(* IEC 61131-3 sources: axsharp/src/ix.compiler/tests/Ix.Compiler.CsTests/samples/units/src, 32 files *)

(* ---- compileromitsattribute.st ---- *)
NAMESPACE CompilerOmmits
    CLASS ClassWithArrays
        VAR PUBLIC
            {#ix-attr:[CompilerOmitsAttribute()]}
            _must_be_omitted_everywhere : Complex;
            {#ix-attr:[CompilerOmitsAttribute("Onliner")]}
            _must_be_omitted_in_onliner : Complex;
            {#ix-attr:[CompilerOmitsAttribute("POCO")]}
             _must_be_omitted_in_poco : Complex;
            _primitive  : ARRAY[0..10] OF BYTE;
        END_VAR

    END_CLASS

    CLASS PUBLIC Complex
        VAR PUBLIC
            HelloString : STRING;
            Id : ULINT;
        END_VAR
    END_CLASS
END_NAMESPACE

NAMESPACE Enums
    CLASS ClassWithEnums
        VAR PUBLIC
            colors : Colors;
            NamedValuesColors : NamedValuesColors;
        END_VAR

    END_CLASS

    TYPE
        Colors : (Red, Green, Blue) := Red;
    END_TYPE

    TYPE
        NamedValuesColors : STRING (Red := '1', Green := '2', Blue := '3') := Red;
    END_TYPE

END_NAMESPACE

NAMESPACE misc
    CLASS PUBLIC VariousMembers
        VAR PUBLIC
            _SomeClass : SomeClass;
            _Motor : Motor;
        END_VAR
    END_CLASS

    CLASS SomeClass
        VAR PUBLIC
            SomeClassVariable : STRING;
        END_VAR
    END_CLASS

    TYPE
        Motor : STRUCT
            isRunning : BOOL;
        END_STRUCT;
        Vehicle : STRUCT
            m : Motor;
            displacement : INT;
        END_STRUCT;
    END_TYPE
END_NAMESPACE

NAMESPACE UnknownArraysShouldNotBeTraspiled
    CLASS ClassWithArrays
        VAR PUBLIC
            _complexKnown : ARRAY[0..10] OF Complex;
            _complexUnknown : ARRAY [0..10] OF ComplexUnknown;
            _primitive  : ARRAY[0..10] OF BYTE;
        END_VAR

    END_CLASS

    CLASS PUBLIC Complex
        VAR PUBLIC
            HelloString : STRING;
            Id : ULINT;
        END_VAR
    END_CLASS
END_NAMESPACE

(* ---- enum_simple.st ---- *)
TYPE
    Colors : (Red, Green, Blue) := Red;
END_TYPE

(* ---- misc.st ---- *)
NAMESPACE Enums
    CLASS ClassWithEnums
        VAR PUBLIC
            colors : Colors;
            NamedValuesColors : NamedValuesColors;
        END_VAR

    END_CLASS

    TYPE
        Colors : (Red, Green, Blue) := Red;
    END_TYPE

    TYPE
        NamedValuesColors : STRING (Red := '1', Green := '2', Blue := '3') := Red;
    END_TYPE

END_NAMESPACE

NAMESPACE misc
    CLASS PUBLIC VariousMembers
        VAR PUBLIC
            _SomeClass : SomeClass;
            _Motor : Motor;
        END_VAR
    END_CLASS

    CLASS SomeClass
        VAR PUBLIC
            SomeClassVariable : STRING;
        END_VAR
    END_CLASS

    TYPE
        Motor : STRUCT
            isRunning : BOOL;
        END_STRUCT;
        Vehicle : STRUCT
            m : Motor;
            displacement : INT;
        END_STRUCT;
    END_TYPE
END_NAMESPACE

NAMESPACE UnknownArraysShouldNotBeTraspiled
    CLASS ClassWithArrays
        VAR PUBLIC
            _complexKnown : ARRAY[0..10] OF Complex;
            _complexUnknown : ARRAY [0..10] OF ComplexUnknown;
            _primitive  : ARRAY[0..10] OF BYTE;
        END_VAR

    END_CLASS

    CLASS PUBLIC Complex
        VAR PUBLIC
            HelloString : STRING;
            Id : ULINT;
        END_VAR
    END_CLASS
END_NAMESPACE

(* ---- struct_simple.st ---- *)
TYPE
    Motor : STRUCT
        isRunning : BOOL;
    END_STRUCT;
    Vehicle : STRUCT
        m : Motor;
        displacement : INT;
    END_STRUCT;
END_TYPE

(* ---- type_named_values.st ---- *)
NAMESPACE NamedValuesNamespace
    TYPE
        LightColors : INT (
            LRED := 12,
            LGREEN := 14,
            LBLUE := 23
        );
    END_TYPE

    CLASS PUBLIC using_type_named_values
        VAR PUBLIC
            LColors : LightColors;
        END_VAR
    END_CLASS
END_NAMESPACE

(* ---- type_named_values_literals.st ---- *)
NAMESPACE Simatic.Ax.StateFramework
    TYPE
        StateControllerStatus : WORD (
            STATUS_NO_ERR := WORD#16#7000,
            STATUS_IS_RUNNING := WORD#16#7001,
            STATUS_STATE_CHANGED := WORD#16#7002,
            STATUS_NO_INITIALSTATE := WORD#16#8100,
            STATUS_NO_NEXTSTATE := WORD#16#8101
        ) := STATUS_NO_ERR;
    END_TYPE

    CLASS PUBLIC using_type_named_values
        VAR PUBLIC
            LColors : StateControllerStatus;
        END_VAR
    END_CLASS
END_NAMESPACE

(* ---- type_with_enum.st ---- *)
NAMESPACE Simatic.Ax.StateFramework
    INTERFACE IGuard

        METHOD Check : BOOL
        END_METHOD

        METHOD Reset
        END_METHOD

    END_INTERFACE
END_NAMESPACE

NAMESPACE Simatic.Ax.StateFramework

    /// Condition
    /// GT: Greater than compareValue
    /// EQ: Equal to compareValue
    /// LT: Less than compareValue
    /// NE: Is not equal to compareValue
    /// GE: Greater or equal to compareValue
    /// LE: Less or equal to compareValue
    TYPE
        Condition : (GT, EQ, LT, NE, GE, LE);
    END_TYPE

    CLASS CompareGuardLint IMPLEMENTS IGuard
        VAR PUBLIC
            Value : REF_TO LINT;
            CompareToValue : LINT;
            Condition : Condition;
        END_VAR

        METHOD PUBLIC Config
            VAR_INPUT
                countValue : REF_TO LINT;
                compareValue : LINT;
                compareCondition : Condition;
            END_VAR
            Value := countValue;
            CompareToValue := compareValue;
            Condition := compareCondition;
        END_METHOD

        // ---------------- IMPLEMENT IGuard---------------------------
        METHOD PUBLIC Check : BOOL

            CASE Condition OF
                Condition#GT : Check := Value^ > CompareToValue;
                Condition#EQ : Check := Value^ = CompareToValue;
                Condition#LT : Check := Value^ < CompareToValue;
                Condition#GE : Check := Value^ >= CompareToValue;
                Condition#LE : Check := Value^ <= CompareToValue;
            END_CASE
            ;

        END_METHOD

        METHOD PUBLIC Reset
            ;
        END_METHOD
        // ---------------- END IMPLEMENT IGuard---------------------------

    END_CLASS
END_NAMESPACE

(* ---- types_with_name_attributes.st ---- *)
NAMESPACE TypeWithNameAttributes
    TYPE
        {#ix-attr:[Container(Layout.Wrap)]}
        Motor : STRUCT
            isRunning : BOOL;
        END_STRUCT;
        Vehicle : STRUCT
            m : Motor;
            displacement : INT;
        END_STRUCT;
    END_TYPE

    {#ix-prop:public string AttributeName}
    CLASS NoAccessModifierClass
        VAR PUBLIC
            SomeClassVariable : STRING;
        END_VAR
    END_CLASS
END_NAMESPACE

(* ---- class_extends_and_implements.st ---- *)
CLASS PUBLIC ExtendsAndImplements EXTENDS ExtendeeExtendsAndImplements IMPLEMENTS IImplementation1, IImplementation2

END_CLASS

CLASS PUBLIC ExtendeeExtendsAndImplements

END_CLASS

INTERFACE PUBLIC IImplementation1 END_INTERFACE
INTERFACE PUBLIC IImplementation2 END_INTERFACE

(* ---- class_implements.st ---- *)
CLASS PUBLIC _NULL_CONTEXT IMPLEMENTS IContext

END_CLASS

INTERFACE PUBLIC IContext

END_INTERFACE

(* ---- class_implements_multiple.st ---- *)
CLASS PUBLIC _NULL_CONTEXT_MULTIPLE IMPLEMENTS IContext_Multiple, IObject_Multiple

END_CLASS

INTERFACE PUBLIC IContext_Multiple

END_INTERFACE

INTERFACE PUBLIC IObject_Multiple

END_INTERFACE

(* ---- file_with_unsupported.st ---- *)
NAMESPACE Unsupported
  FUNCTION SomeFunction : INT
    ;
  END_FUNCTION
END_NAMESPACE

(* ---- array_declaration.st ---- *)
NAMESPACE ArrayDeclarationSimpleNamespace
    CLASS array_declaration_class
        VAR PUBLIC
            primitive : ARRAY[1..100] OF INT;
            complex : ARRAY[1..100] OF some_complex_type;
        END_VAR
    END_CLASS

    CLASS some_complex_type
        VAR

        END_VAR

    END_CLASS

END_NAMESPACE

(* ---- class_all_primitives.st ---- *)
CLASS class_all_primitives
    VAR PUBLIC
        myBOOL	        :       BOOL	      ;
        myBYTE	        :       BYTE	      ;
        myWORD	        :       WORD	      ;
        myDWORD	        :       DWORD	      ;
        myLWORD	        :       LWORD	      ;
        mySINT	        :       SINT	      ;
        myINT	        :       INT	          ;
        myDINT	        :       DINT	      ;
        myLINT	        :       LINT	      ;
        myUSINT	        :       USINT	      ;
        myUINT	        :       UINT	      ;
        myUDINT	        :       UDINT	      ;
        myULINT	        :       ULINT	      ;
        myREAL	        :       REAL	      ;
        myLREAL	        :       LREAL	      ;
        myTIME	        :       TIME	      ;
        myLTIME	        :       LTIME	      ;
        myDATE	        :       DATE	      ;
     //   myLDATE	        :       LDATE	      ;
        myTIME_OF_DAY	:       TIME_OF_DAY	  ;
     //   myLTIME_OF_DAY	:       LTIME_OF_DAY  ;
        myDATE_AND_TIME  :      DATE_AND_TIME ;
     //   myLDATE_AND_TIME :      LDATE_AND_TIME;
     //   myCHAR	        :       CHAR	      ;
     //   myWCHAR	        :       WCHAR	      ;
        mySTRING	        :   STRING	      ;
        myWSTRING	    :       WSTRING	      ;
    END_VAR
END_CLASS

(* ---- class_extended_by_known_type.st ---- *)
USING Simatic.Ax.Stateframework;
USING Simatic.Ax.StatePattern;

NAMESPACE Simatic.Ax.StateFramework
    CLASS State1Transition EXTENDS AbstractState

        METHOD PUBLIC OVERRIDE OnEntry
            ;
        END_METHOD

        METHOD PUBLIC OVERRIDE OnExit
            ;
        END_METHOD

        METHOD PUBLIC OVERRIDE Action
            ;
        END_METHOD

    END_CLASS

END_NAMESPACE

NAMESPACE Simatic.Ax.StateFramework
    CLASS ABSTRACT AbstractState IMPLEMENTS IState, IStateMuteable

        VAR PUBLIC
            Transition1 : ITransition;
            StateID : INT;
            StateName : String;
        END_VAR

        VAR PROTECTED
             _actualStatus : StateStatus;
        END_VAR

        // METHOD PUBLIC ABSTRACT OnEntry
        // END_METHOD
        METHOD PUBLIC OnEntry
            _actualStatus := StateStatus#Active;
        END_METHOD

        METHOD PUBLIC ABSTRACT OnExit
        END_METHOD

        METHOD PUBLIC ABSTRACT Action
        END_METHOD

        METHOD PUBLIC GetTransition : ITransition
            VAR_INPUT
                pos : UINT;
            END_VAR
            IF (THIS.TransitionCount() = pos + UINT#1) THEN
                GetTransition := transition1;
            ELSE
                GetTransition := NULL;
            END_IF;
        END_METHOD

        METHOD PUBLIC TransitionCount : UINT
            IF (transition1 <> NULL) THEN
                TransitionCount := UINT#1;
            ELSE
                TransitionCount := UINT#0;
            END_IF;
        END_METHOD

        METHOD PUBLIC GetStateID : INT
            GetStateID := StateID;
        END_METHOD

        METHOD PUBLIC FINAL GetStateName : STRING
            GetStateName := StateName;
        END_METHOD

        METHOD PUBLIC FINAL GetStatus : StateStatus
            GetStatus := _actualStatus;
        END_METHOD

        METHOD PUBLIC FINAL SetStatus
            VAR_INPUT
                status : StateStatus;
            END_VAR
            _actualStatus := status;
        END_METHOD
    END_CLASS
END_NAMESPACE

(* ---- class_extends.st ---- *)
CLASS PUBLIC Extended EXTENDS Extendee

END_CLASS

CLASS PUBLIC Extendee

END_CLASS

(* ---- class_internal.st ---- *)
CLASS INTERNAL ClassWithComplexTypes

END_CLASS

(* ---- class_no_access_modifier.st ---- *)
CLASS NoAccessModifierClass

END_CLASS

(* ---- class_with_complex_members.st ---- *)
NAMESPACE ClassWithComplexTypesNamespace
    CLASS PUBLIC ClassWithComplexTypes
        VAR PUBLIC
           myComplexType : ComplexType1;
        END_VAR
    END_CLASS

    CLASS PUBLIC ComplexType1

    END_CLASS
END_NAMESPACE

(* ---- class_with_non_public_members.st ---- *)
NAMESPACE ClassWithNonTraspilableMemberssNamespace
    CLASS PUBLIC ClassWithNonTraspilableMembers
        VAR PUBLIC
           myComplexType : ComplexType1;
        END_VAR

        VAR
           myComplexType1 : ComplexType1;
           myBooool : BOOL;
        END_VAR

        VAR
           myComplexType2 : ComplexType1;
           myBooool1 : BOOL;
        END_VAR
    END_CLASS

    CLASS PUBLIC ComplexType1

    END_CLASS
END_NAMESPACE

(* ---- class_with_pragmas.st ---- *)
NAMESPACE ClassWithPragmasNamespace
    {#ix-attr:[Container(Layout.Stack)]}
    CLASS PUBLIC  ClassWithPragmas
        VAR PUBLIC
           {#ix-attr:[Container(Layout.Wrap)]}
           myComplexType : ComplexType1;
        END_VAR
    END_CLASS

    CLASS PUBLIC ComplexType1

    END_CLASS
END_NAMESPACE

(* ---- class_with_primitive_members.st ---- *)
NAMESPACE ClassWithPrimitiveTypesNamespace
    CLASS PUBLIC ClassWithPrimitiveTypes
        VAR PUBLIC
           myBOOL	        :       BOOL	      ;
           myBYTE	        :       BYTE	      ;
           myWORD	        :       WORD	      ;
           myDWORD	        :       DWORD	      ;
           myLWORD	        :       LWORD	      ;
           mySINT	        :       SINT	      ;
           myINT	        :       INT	          ;
           myDINT	        :       DINT	      ;
           myLINT	        :       LINT	      ;
           myUSINT	        :       USINT	      ;
           myUINT	        :       UINT	      ;
           myUDINT	        :       UDINT	      ;
           myULINT	        :       ULINT	      ;
           myREAL	        :       REAL	      ;
           myLREAL	        :       LREAL	      ;
           myTIME	        :       TIME	      ;
           myLTIME	        :       LTIME	      ;
           myDATE	        :       DATE	      ;
           myLDATE	        :       LDATE	      ;
           myTIME_OF_DAY	:       TIME_OF_DAY	  ;
           myLTIME_OF_DAY	:       LTIME_OF_DAY  ;
           myDATE_AND_TIME  :       DATE_AND_TIME ;
           myLDATE_AND_TIME :       LDATE_AND_TIME;
           myCHAR	        :       CHAR	      ;
           myWCHAR	        :       WCHAR	      ;
           mySTRING	        :       STRING	      ;
           myWSTRING	    :       WSTRING	      ;
        END_VAR
    END_CLASS
END_NAMESPACE

(* ---- class_with_using_directives.st ---- *)
CLASS INTERNAL ClassWithUsingDirectives
    USING SimpleFirstLevelNamespace, SimpleQualifiedNamespace.Qualified;
    USING HelloLevelOne.HelloLevelTwo;
    USING InexistingNamespace;
END_CLASS

NAMESPACE SimpleFirstLevelNamespace

END_NAMESPACE

NAMESPACE SimpleQualifiedNamespace.Qualified

END_NAMESPACE

NAMESPACE HelloLevelOne
    NAMESPACE HelloLevelTwo
    END_NAMESPACE
END_NAMESPACE

(* ---- configuration.st ---- *)
CONFIGURATION MyConfiguration
    TASK Main(Interval := T#1000ms, Priority := 1);
    PROGRAM P1 WITH Main: MyProgram;

    VAR_GLOBAL
        Complex : ComplexForConfig;
        myBOOL	        :       BOOL	      ;
        myBYTE	        :       BYTE	      ;
        myWORD	        :       WORD	      ;
        myDWORD	        :       DWORD	      ;
        myLWORD	        :       LWORD	      ;
        mySINT	        :       SINT	      ;
        myINT	        :       INT	          ;
        myDINT	        :       DINT	      ;
        myLINT	        :       LINT	      ;
        myUSINT	        :       USINT	      ;
        myUINT	        :       UINT	      ;
        myUDINT	        :       UDINT	      ;
        myULINT	        :       ULINT	      ;
        myREAL	        :       REAL	      ;
        myLREAL	        :       LREAL	      ;
        myTIME	        :       TIME	      ;
        myLTIME	        :       LTIME	      ;
        myDATE	        :       DATE	      ;
        myLDATE	        :       LDATE	      ;
        myTIME_OF_DAY	:       TIME_OF_DAY	  ;
        myLTIME_OF_DAY	:       LTIME_OF_DAY  ;
        myDATE_AND_TIME  :       DATE_AND_TIME ;
        myLDATE_AND_TIME :       LDATE_AND_TIME;
        myCHAR	        :       CHAR	      ;
        myWCHAR	        :       WCHAR	      ;
        mySTRING	        :       STRING	      ;
        myWSTRING	    :       WSTRING	      ;

        {#ix-attr:[ReadOnce()]}
        myWSTRING_readOnce	    :       WSTRING	      ;
        {#ix-attr:[ReadOnly()]}
        myWSTRING_readOnly	    :       WSTRING	      ;
        {#ix-attr:[ReadOnce()]}
        cReadOnce           : ComplexForConfig;
        {#ix-attr:[ReadOnly()]}
        cReadOnly           : ComplexForConfig;
        Colorss : Colorss;
        Colorsss : Colorsss;

        {#ix-attr:[CompilerOmitsAttribute()]}
        _must_be_omitted_everywhere : BOOL;
        {#ix-attr:[CompilerOmitsAttribute("Onliner")]}
        _must_be_omitted_in_onliner : BOOL;
        {#ix-attr:[CompilerOmitsAttribute("POCO")]}
         _must_be_omitted_in_poco : BOOL;
    END_VAR
END_CONFIGURATION

CLASS PUBLIC ComplexForConfig
    VAR PUBLIC
        myBOOL	        :       BOOL	      ;
        myBYTE	        :       BYTE	      ;
        myWORD	        :       WORD	      ;
        myDWORD	        :       DWORD	      ;
        myLWORD	        :       LWORD	      ;
        mySINT	        :       SINT	      ;
        myINT	        :       INT	          ;
        myDINT	        :       DINT	      ;
        myLINT	        :       LINT	      ;
        myUSINT	        :       USINT	      ;
        myUINT	        :       UINT	      ;
        myUDINT	        :       UDINT	      ;
        myULINT	        :       ULINT	      ;
        myREAL	        :       REAL	      ;
        myLREAL	        :       LREAL	      ;
        myTIME	        :       TIME	      ;
        myLTIME	        :       LTIME	      ;
        myDATE	        :       DATE	      ;
        myLDATE	        :       LDATE	      ;
        myTIME_OF_DAY	:       TIME_OF_DAY	  ;
        myLTIME_OF_DAY	:       LTIME_OF_DAY  ;
        myDATE_AND_TIME  :       DATE_AND_TIME ;
        myLDATE_AND_TIME :       LDATE_AND_TIME;
        myCHAR	        :       CHAR	      ;
        myWCHAR	        :       WCHAR	      ;
        mySTRING	        :       STRING	      ;
        myWSTRING	    :       WSTRING	      ;
    END_VAR
END_CLASS

TYPE
    Colorss : (Red, Green, Blue) := Red;
END_TYPE

TYPE
    Colorsss : ULINT (Red := ULINT#1, Green := ULINT#2, Blue := ULINT#3) := Red;
END_TYPE

(* ---- makereadonce.st ---- *)
NAMESPACE makereadonce
    CLASS PUBLIC MembersWithMakeReadOnce
        VAR PUBLIC
            {#ix-attr:[ReadOnce()]}
            makeReadOnceMember : STRING;
            someOtherMember : STRING;

            {#ix-attr:[ReadOnce()]}
            makeReadComplexMember : ComplexMember;
            someotherComplexMember : ComplexMember;
        END_VAR
    END_CLASS

    CLASS PUBLIC ComplexMember
        VAR PUBLIC
            someMember : STRING;
            someOtherMember : STRING;
        END_VAR
    END_CLASS
END_NAMESPACE

(* ---- makereadonly.st ---- *)
NAMESPACE makereadonly
    CLASS PUBLIC MembersWithMakeReadOnly
        VAR PUBLIC
            {#ix-attr:[ReadOnly()]}
            makeReadOnceMember : STRING;
            someOtherMember : STRING;

            {#ix-attr:[ReadOnly()]}
            makeReadComplexMember : ComplexMember;
            someotherComplexMember : ComplexMember;
        END_VAR
    END_CLASS

    CLASS PUBLIC ComplexMember
        VAR PUBLIC
            someMember : STRING;
            someOtherMember : STRING;
        END_VAR
    END_CLASS
END_NAMESPACE

(* ---- ref_to_simple.st ---- *)
NAMESPACE RefToSimple
    CLASS ref_to_simple
        VAR PUBLIC
            a : REF_TO INT;
            b : REF_TO referenced;
        END_VAR
    END_CLASS

    CLASS referenced
        VAR PUBLIC
            b : INT;
        END_VAR
    END_CLASS
END_NAMESPACE

(* ---- simple_empty_class.st ---- *)
CLASS PUBLIC simple_class
END_CLASS

(* ---- simple_empty_class_within_namespace.st ---- *)
NAMESPACE sampleNamespace
    CLASS PUBLIC simple_empty_class_within_namespace
    END_CLASS
END_NAMESPACE

(* ---- types_with_property_attributes.st ---- *)
NAMESPACE TypesWithPropertyAttributes
    {#ix-prop:public string Description}
    {#ix-set:Description = "Some added property name value"}
    CLASS SomeAddedProperties
        VAR PUBLIC
            {#ix-set:AttributeName = "Pocitadlo"}
            Counter : INT;
        END_VAR
    END_CLASS
END_NAMESPACE

(* ---- file_with_usings.st ---- *)
USING FileWithUsingsSimpleFirstLevelNamespace;
USING FileWithUsingsSimpleQualifiedNamespace.Qualified;
USING FileWithUsingsHelloLevelOne.FileWithUsingsHelloLevelTwo;

NAMESPACE FileWithUsingsSimpleFirstLevelNamespace

END_NAMESPACE

NAMESPACE FileWithUsingsSimpleQualifiedNamespace.Qualified

END_NAMESPACE

NAMESPACE FileWithUsingsHelloLevelOne
    NAMESPACE FileWithUsingsHelloLevelTwo
    END_NAMESPACE
END_NAMESPACE

(* ---- program.st ---- *)
PROGRAM MyProgram
    VAR_EXTERNAL

    END_VAR

    VAR

    END_VAR

    VAR_TEMP

    END_VAR

    // code here
    ;
END_PROGRAM
